// FB EDM state codes.
{attribute 'qualified_only'}
{attribute 'to_string'}
TYPE
E_SafeEdmState :
(
    Undefined := 0,
    Stop := 2,
    Error := 4,
    Reset := 5,
    MonOff := 14,
    MonOn := 15
) BYTE;
END_TYPE

(* stored: Version 1.1.0.1
   DUT E_SafeEdmState: Id {dc1d1a43-a154-599b-a2b5-f267c93c1dad} *)
